(* IEC 61131-3 sources: plc-vscode/tests/st/all/rusty/tests/lit/multi/cross_unit_dependency_resolution, 1 file *)

(* ---- main.st ---- *)
FUNCTION test_function : BOOL
VAR_INPUT
    input_data : struct_array;
END_VAR
VAR_IN_OUT
    output_data : struct_array;
END_VAR
    test_function := TRUE;
END_FUNCTION

FUNCTION main : DINT
VAR
    // Array of typedef of struct
    my_struct_arr : struct_array;

    // Array of typedef of array
    nested_arr : ARRAY[0..1] OF int_array;

    // Pointer to typedef of struct
    struct_pointer : struct_ptr;

    // Pointer to typedef of array
    array_pointer : array_ptr;

    // Complex container
    container : container_struct;

    // Multi-dimensional
    matrix : matrix_type;

    // Deep typedef chain
    deep_var : level2_typedef;

    // Array of typedef of struct of array
    complex_nested : complex_nested_array;

    // Typedef struct of struct
    typedef_nested : typedef_nested_struct;

    // Struct of struct
    direct_nested : direct_nested_struct;
END_VAR
    my_struct_arr[0].x := 1337;
    my_struct_arr[0].y := 3.14;

    deep_var.x := 7331;
    deep_var.y := 2.71;

    container.arr_field[0].x := 9001;
    container.status := status_enum#RUNNING;
    container.percent := 75;

    matrix[0][0] := 1.23;
    matrix[1][1] := 4.56;

    test_function(my_struct_arr, my_struct_arr);

    complex_nested[0].values[0] := 42;
    complex_nested[0].count := 84;

    typedef_nested.outer_field.x := 1000;
    typedef_nested.outer_field.y := 2.5;
    typedef_nested.inner.values[0] := 123;

    direct_nested.outer_field.x := 2000;
    direct_nested.outer_field.y := 5.0;
    direct_nested.inner.values[1] := 456;

    printf('%d$N', my_struct_arr[0].x);     // CHECK: 1337
    printf('%.2f$N', my_struct_arr[0].y);   // CHECK: 3.14
    printf('%d$N', deep_var.x);             // CHECK: 7331
    printf('%.2f$N', deep_var.y);           // CHECK: 2.71
    printf('%d$N', container.arr_field[0].x); // CHECK: 9001
    printf('%d$N', container.status);       // CHECK: 1
    printf('%d$N', container.percent);      // CHECK: 75
    printf('%.2f$N', matrix[0][0]);         // CHECK: 1.23
    printf('%.2f$N', matrix[1][1]);         // CHECK: 4.56
    printf('%d$N', complex_nested[0].values[0]); // CHECK: 42
    printf('%d$N', complex_nested[0].count); // CHECK: 84
    printf('%d$N', typedef_nested.outer_field.x); // CHECK: 1000
    printf('%.1f$N', typedef_nested.outer_field.y); // CHECK: 2.5
    printf('%d$N', typedef_nested.inner.values[0]); // CHECK: 123
    printf('%d$N', direct_nested.outer_field.x); // CHECK: 2000
    printf('%.1f$N', direct_nested.outer_field.y); // CHECK: 5.0
    printf('%d$N', direct_nested.inner.values[1]); // CHECK: 456

    main := 0;
END_FUNCTION
